RoboDK station: weldcell.rdk

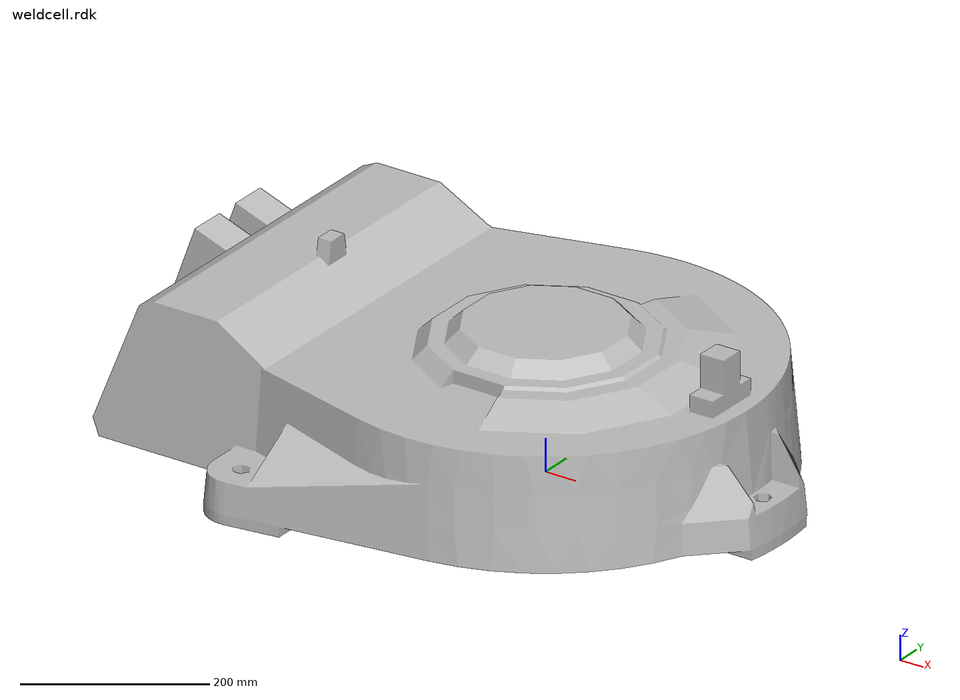
[picture v0: the station drawn from its stored meshes, robots at their saved joint values, targets as dots, program paths as lines]
Station weldcell (saved by RoboDK 6.2.0). Poses are relative to the parent item; angles as X-Y-Z fixed-axis rotations.
  - frame ABB IRB 2400/16 Base at (0, 0, 0) mm
    - robot ABB IRB 2400/16: 6 axes, payload 16 kg, reach 1550 mm, repeatability 0.03 mm, weight 380 kg
        joint limits [-180, -100, -60, -200, -120, -400] to [180, 110, 65, 200, 120, 400]; home [0, 0, 0, 0, 0, 0]; saved at [0, 0, 0, 0, 0, 0]
